Fanuc KAREL source: KB00133.KL

PROGRAM KB00133
%NOLOCKGROUP
%ENVIRONMENT REGOPE
VAR
  P1: INTEGER
  P2: INTEGER
  P3: INTEGER
  P4: INTEGER
  P5: INTEGER
BEGIN
  P1 = 1
  P2 = 1
  P3 = 1
  P4 = 1
  P5 = 1
  POS_REG_TYPE(P1, P2, P3, P4, P5)
END KB00133
